(* IEC 61131-3 sources: Pirate/PLC/DUT, 3 files *)

(* ---- ST_AreteZone.st ---- *)
TYPE ST_AreteZone :
STRUCT
    NoeudA : UINT; // indice dans le tableau des noeuds de la zone
    NoeudB : UINT; // indice dans le tableau des noeuds de la zone
    EquipementIndex : INT; // -1 pour une liaison permanente, sinon indice equipement
END_STRUCT
END_TYPE

(* ---- ST_Equipement.st ---- *)
TYPE ST_Equipement :
STRUCT
    Id : UINT; // identifiant unique dans la zone (1..80)
    Ferme : BOOL; // commande ou position simulee
    Defaut : BOOL; // indisponibilite : coupe la conduction
    Asservi : BOOL; // TRUE si l'equipement est soumis a un asservissement (non implemente)
    Conducteur : BOOL; // resultat calcule par FB_Zone
END_STRUCT
END_TYPE

(* ---- ST_Noeud.st ---- *)
TYPE ST_Noeud :
STRUCT
    IdZone : UINT; // identifiant metier (1..57)
    SousTension : BOOL; // resultat du parcours BFS
END_STRUCT
END_TYPE
